FUNCTION_BLOCK DataType
  (* Standard: 61499-1; Description: Copyright (c) 2026 Martin Erich Jobst This program and the accompanying materials are made available under the terms of the Eclipse Public License 2.0 which is available at https://www.eclipse.org/legal/epl-2.0/ SPDX-License-Identifier: EPL-2.0 *)
  (* Version 1.0, 2026-11-18, Martin Jobst *)
  PACKAGE lib::ConfigurableFB;
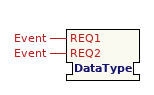
  EVENT_INPUT
    REQ1;
    REQ2;
  END_EVENT
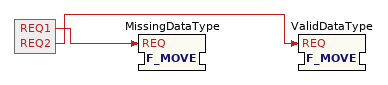
  FBS
    MissingDataType : iec61131::selection::F_MOVE; {SET_ATTRIBUTE(DataType, MissingDataType)}
    ValidDataType : iec61131::selection::F_MOVE; {SET_ATTRIBUTE(DataType, DINT)}
  END_FBS
  EVENT_CONNECTIONS
    REQ1 TO MissingDataType.REQ;
    REQ2 TO ValidDataType.REQ;
  END_CONNECTIONS
END_FUNCTION_BLOCK
